(*
SPDX-FileCopyrightText: © 2026 Oleksandr Tiutyk <trofimich@gmail.com>
SPDX-License-Identifier: MIT
License: https://opensource.org/license/mit
*)

(*!
<summary>Records automatic execution error recoveries for analog input tests.</summary>
<description>Uses the inherited analog input constructor, processing, and error handling.</description>
*)
{attribute 'no_explicit_call' := 'do not call this function block directly'}
FUNCTION_BLOCK FINAL AnalogInputRecoveryProbe EXTENDS TOF_Devices_IO.AnalogInput
VAR
	_RecoveryCalls : UDINT;
END_VAR

(*!
<summary>Counts the recovery callback issued by Execute().</summary>
*)
METHOD PROTECTED OnRecover
_RecoveryCalls := _RecoveryCalls + UDINT#1;
END_METHOD

(*!
<summary>Gets the number of recovery callbacks received by this instance.</summary>
*)
PROPERTY RecoveryCalls : UDINT
GET
RecoveryCalls := _RecoveryCalls;
END_GET
END_PROPERTY

END_FUNCTION_BLOCK

(* stored: Version 1.1.0.1
   POU AnalogInputRecoveryProbe: Id {651d0ebf-17f4-4020-a80c-5bdcb4d1cb93}, SpecialFunc None
   Method OnRecover: Id {df5058c8-ef9e-4ead-b573-aadfe29f3931}
   Property RecoveryCalls: Id {8dbae345-0861-4232-b263-6e426b022de5}
   Get Get: Id {c278a49e-d1bc-405a-aa6b-7d4e98e7ab0c} *)
